Fanuc KAREL source: kt00340.KL

-- PROVISIONAL review KL for V1013-1; original PC SHA256 10e6b39082c183af295b2ccaf7f07e0c248c9776f3b57bd57f3177b5a2cbad0a
-- Incomplete behavior may be omitted. Consult companion uncertainty JSON. Do not deploy.
PROGRAM KT00340
%NOLOCKGROUP
VAR
  R2 : REAL
  OUT : BOOLEAN
-- UNRESOLVED_DECL Y1 type=002018
BEGIN
  -- UNRESOLVED_PC offsets 5-19; opcodes 2E,22,9D,33,B2
  -- UNRESOLVED_PC offsets 24-35; opcodes 2E,23
  -- UNRESOLVED_PC offsets 40-65; opcodes 22,9D,33,B1,21,29,64,29,6F,23
  -- UNRESOLVED_PC offsets 70-74; opcodes 7F
END KT00340
